// TIA Portal V21 export
// export: Created 2026-10-12T11:32:17.3982992Z, ExportSetting WithDefaults, DisplayName Totally Integrated Automation Portal, DisplayVersion V21, DisplayName STEP 7 Professional, DisplayVersion V21, DisplayName STEP 7 Safety, DisplayVersion V21, DisplayName Tech WebApplication, DisplayVersion V21, DisplayName WinCC Basic/Comfort/Advanced, DisplayVersion V21, DisplayName WinCC Unified, DisplayVersion V21
VAR_GLOBAL   // PLC tag table "DO"
   "DO_CONVEYOR FWD ON" AT %Q0.0 : Bool;
   "DO_CONVEYOR REV ON" AT %Q0.1 : Bool;
   "DO_FAULT RESET" AT %Q0.2 : Bool;
   "DO_TL GREEN" AT %Q0.3 : Bool;
   "DO_TL RED" AT %Q0.4 : Bool;
   "DO_TL AMBER" AT %Q0.5 : Bool;
   "DO_SPARE Q0.6" AT %Q0.6 : Bool;
   "DO_SPARE Q0.7" AT %Q0.7 : Bool;
   "DO_SPARE Q1.0" AT %Q1.0 : Bool;
   "DO_SPARE Q1.1" AT %Q1.1 : Bool;
END_VAR
